Staubli VAL3: search_traj.pgx

program search_traj(bool& x_bFounded, string& x_sSessionName, num x_nSession)
  local string l_sEmpty
  local num i
  local num l_nSession
  local bool l_bOk
begin
  // init
  x_bFounded=false
  x_sSessionName=""
  //
  // get the list
  //
  l_sEmpty=""
  call trajectory:getTrajList(sSessionList)
  //
  // search the program from a number:
  //
  // "number+space+name"
  //
  // 01 MyPart
  // 10 YourPart
  //
  for i=0 to size(sSessionList)-1
    if sSessionList[i]!=""
      // convert the string "00 name" into a num
      toNum(sSessionList[i],l_nSession,l_bOk)
      if l_bOk and l_nSession==x_nSession
        x_sSessionName=sSessionList[i]
        x_bFounded=true
        // exit
        i=size(sSessionList)-1
      endIf
    endIf
  endFor
end
